Staubli VAL3: init.pgx

public program init()
begin
  //init all
  bIsSaving=false
  call resetAlarm()
  bAlarmAck=false
  bGOTO=false
  bIsCycle=false
  bIsEstop=false
  bIsHome=false
  bIsReady=false
  bReloadIO=false
  bSimulate=false
  bSimulate=false
  _bHeavyAlarm=false
  bQuitApp=false
  nCycleCmd=0
  nCycleMoveID=0
  nFrameIndex=0
  nHeavyAlarmLev=0
  nHMIcmd=0
  nPLCcmd=0
  nToolIndex=0
  _nAlarmIndex=0
  _nAvgCapacity=0
  _nBestCapacity=0
  _nCapacity=0
  _nCTIndex=0
  _nCycleTime=0
  _nOmacStat=9

  sPageUsing=""
  sTrajStatus=""
  sLstTrajStatus=""
  _sRobotStatus=""
  sLstRobStatus=""
  sIOStatus=""
  sLstIOStatus=""

end
